// TIA Portal V19 export
DATA_BLOCK "GenralDB"   // DB18
{ S7_Optimized_Access := 'TRUE' }
// stored: MemoryReserve 100
   VAR
      Solvent_Addition_Running_1 : Bool;
      NBL_Addition_Running_1 : Bool;
   END_VAR
BEGIN
END_DATA_BLOCK
